(* IEC 61131-3 sources: Jog-the-Robot/plc-for-usb, 2 files *)

(* ---- Main.st ---- *)
(*********************************************************************************
 * Copyright: B&R Industrial Automation GmbH
 * Author:    huebnern
 * Created:   January 23, 2020/8:20 AM
 * Edited:    October 26, 2026 - phone jog, power and home via ESP32 (action RemoteJog)
 *********************************************************************************)
//Main control of the system
PROGRAM _INIT

	//Init Status error
	MainPar.VisuPars.InError 	:= FALSE;
	MainPar.VisuPars.NotInError	:= TRUE;

	//Init Jog velocity
	JogVelocity 				:= INIT_JOG_VELOCITY;

	//Allow jog (Icmp_Ping task is not used)
	AllowJog := TRUE;

	Teach_Pos[0].Pos.X						:=	240;
	Teach_Pos[0].Pos.Y						:= 	0;
	Teach_Pos[0].Pos.Z						:=	335;
	Teach_Pos[0].Orient.Angle1				:=	0;
	Teach_Pos[0].Orient.Angle2				:=	0;

	Teach_Pos[1].Pos.X := 20.699866696484403;
	Teach_Pos[1].Pos.Y := -16.763507571369498;
	Teach_Pos[1].Pos.Z	:= 680.95033173265676;
	Teach_Pos[1].Orient.Angle1 := -126.89365872204304;
	Teach_Pos[1].Orient.Angle2 := 140.99818452000619;

	Teach_Pos[2].Pos.X := -69.244968642624457;
	Teach_Pos[2].Pos.Y := 56.0771029659347;
	Teach_Pos[2].Pos.Z	:= 672.76899259820129;
	Teach_Pos[2].Orient.Angle1 := -111.97058904528618;
	Teach_Pos[2].Orient.Angle2 := 140.99818452000619;

	Teach_Pos[3].Pos.X := 240;
	Teach_Pos[3].Pos.Y := 0;
	Teach_Pos[3].Pos.Z	:= 335;
	Teach_Pos[3].Orient.Angle1 := 0;
	Teach_Pos[3].Orient.Angle2 := 0;

END_PROGRAM

PROGRAM _CYCLIC
	Aktor := Sensor;
	//Error Reset
	fbMpRobotic5Arm.ErrorReset				:= MainPar.Cmd.ErrorReset;

	//Write status
	StatusMain;

	//Change visualization vars
	VisuDisable;

	//Phone jog via ESP32 (BLE -> Modbus TCP). Must run before the state machine.
	RemoteJog;

	//Power On
	IF MainPar.Cmd.PowerOn THEN
		IF fbMpRobotic5Arm.Info.ReadyToPowerOn AND MainPar.StateMachine = STATE_Disabled THEN
			MainPar.StateMachine 	:= STATE_PowerOn;
		END_IF
	ELSE
		MainPar.StateMachine 		:= STATE_Disabled;
	END_IF

	//---------------------------------------------
	//-------------State Machine-------------------
	//---------------------------------------------
	CASE MainPar.StateMachine OF

		//--------State Disabled-------------------
		STATE_Disabled:

			//Power robot off
			fbMpRobotic5Arm.Power 			:= FALSE;

			//Set PreStateIdent
			MainPar.PreStateIdent 			:= STATE_Disabled;

			//Reset Error as long as the robot is disabled
			MainPar.VisuPars.InError 	:= FALSE;
			MainPar.VisuPars.NotInError	:= TRUE;

		//--------State PowerOn-------------------
		STATE_PowerOn:

			//Power robot on
			fbMpRobotic5Arm.Power 			:= TRUE;

			IF MainPar.Status = Idle THEN
				MainPar.StateMachine 		:= STATE_WaitForHome;
			END_IF

		//--------State WaitForHome-------------------
		STATE_WaitForHome:

			//Set PreStateIdent
			MainPar.PreStateIdent 			:= STATE_WaitForHome;

			//Reset Stop
			IF fbMpRobotic5Arm.Stop THEN
				fbMpRobotic5Arm.Stop 		:= FALSE;
			END_IF

			IF MainPar.Cmd.Home THEN
				MainPar.StateMachine 	:= STATE_Home;
				MainPar.HomingCount		:= NoHoming;
				//Reset command
				MainPar.Cmd.Home 		:= FALSE;
			END_IF

		//--------State Home-------------------
		STATE_Home:

			fbMpRobotic5Arm.Home := TRUE;

			IF MainPar.HomingCount = NoHoming THEN
				ChangeHomingMode := FALSE;
			ELSIF MainPar.HomingCount = DefaultHomingDone THEN
				ChangeHomingMode := TRUE;
			END_IF

			IF EDGEPOS(fbMpRobotic5Arm.IsHomed) THEN
				MainPar.HomingCount 		:= MainPar.HomingCount + 1;
				fbMpRobotic5Arm.Home 		:= FALSE;
			END_IF

			IF MainPar.HomingCount = DirectHomingDone THEN
				MainPar.StateMachine 		:= STATE_Idle;
				fbMpRobotic5Arm.Home 		:= FALSE;
			ELSIF MainPar.Cmd.Stop THEN
				MainPar.StateMachine 		:= STATE_WaitForHome;
				fbMpRobotic5Arm.Stop 		:= TRUE;
				fbMpRobotic5Arm.Home 		:= FALSE;
				//Reset command
				MainPar.Cmd.Stop 			:= FALSE;
			END_IF

		//--------State Idle-------------------
		STATE_Idle:

			//Set PreStateIdent
			MainPar.PreStateIdent 			:= STATE_Idle;

			//Reset Stop
			IF fbMpRobotic5Arm.Stop THEN
				fbMpRobotic5Arm.Stop 		:= FALSE;
			END_IF

			IF MainPar.Cmd.Home THEN
				MainPar.HomingCount			:= NoHoming;
				MainPar.StateMachine 		:= STATE_Home;

			ELSE

				//Change to GCode state in case of visu is currently on the G-Code page
				IF (MainPar.GoToState.GCode) AND EDGEPOS(MainPar.Cmd.Start) THEN
					MainPar.StateMachine 	:= STATE_GCode;
				END_IF

				//Change to Tipping state in case of visu is currently on the Tipping page (or the phone has control)
				IF (MainPar.GoToState.Tipping) AND (JogDirectionSet) THEN
					MainPar.StateMachine 	:= STATE_Tipping;
				END_IF

				//Change to MoveSetPos state in case of visu is currently on the MoveSetPos page
				IF (MainPar.GoToState.MoveSetPos) AND EDGEPOS(MainPar.Cmd.Start) THEN
					MainPar.StateMachine 	:= STATE_MoveSetPos;
				END_IF

			END_IF

		//--------State G-Code-------------------
		STATE_GCode:

			//Start movement
			fbMpRobotic5Arm.MoveProgram 		:= TRUE;

			//Stop movement
			IF MainPar.Cmd.Stop THEN
				fbMpRobotic5Arm.Stop 			:= TRUE;
				fbMpRobotic5Arm.MoveProgram 	:= FALSE;
				MainPar.StateMachine 			:= STATE_Idle;
			ELSIF fbMpRobotic5Arm.MoveDone THEN
				fbMpRobotic5Arm.MoveProgram 	:= FALSE;
				MainPar.StateMachine 			:= STATE_Idle;
			END_IF

		//--------State Tipping-------------------
		STATE_Tipping:

			//Change coordinate system
			ParRobot.CoordSystem 			:= mcACS;

			//Set velocity for chosen axis with action
			Tipping;

			//Call Jog
			IF AllowJog THEN
				fbMpRobotic5Arm.Jog := TRUE;
			ELSE
				fbMpRobotic5Arm.Jog := FALSE;
			END_IF

			IF NOT JogDirectionSet THEN
				MainPar.StateMachine 		:= STATE_Idle;
				fbMpRobotic5Arm.Jog 		:= FALSE;
			END_IF

		//--------State MoveSetPos-------------------
		STATE_MoveSetPos:

			//Change coordinate system
			ParRobot.CoordSystem 				:= mcMCS;

			//Start movement
			IF MainPar.Cmd.MoveIndex THEN
				fbMpRobotic5Arm.MoveDirect 	:= TRUE;
			ELSIF NOT MainPar.Cmd.MoveIndex THEN
				fbMpRobotic5Arm.MoveLinear 	:= TRUE;
			END_IF

			//Stop movement
			IF MainPar.Cmd.Stop THEN
				fbMpRobotic5Arm.Stop 			:= TRUE;
				fbMpRobotic5Arm.MoveDirect 	:= FALSE;
				fbMpRobotic5Arm.MoveLinear 	:= FALSE;
				MainPar.StateMachine 			:= STATE_Idle;
			ELSIF fbMpRobotic5Arm.MoveDone THEN
				fbMpRobotic5Arm.MoveDirect 	:= FALSE;
				fbMpRobotic5Arm.MoveLinear 	:= FALSE;
				MainPar.StateMachine 			:= STATE_Idle;
			END_IF

		//--------State Error-------------------
		STATE_Error:

			//Set output var for visu
			MainPar.VisuPars.InError 		:= TRUE;
			MainPar.VisuPars.NotInError		:= FALSE;

			//Stop movement
			fbMpRobotic5Arm.Stop 			:= TRUE;
			fbMpRobotic5Arm.MoveDirect 	:= FALSE;
			fbMpRobotic5Arm.MoveLinear 	:= FALSE;
			fbMpRobotic5Arm.Jog 			:= FALSE;
			fbMpRobotic5Arm.MoveProgram 	:= FALSE;
			fbMpRobotic5Arm.Home 			:= FALSE;

			//Go out of the error state as soon as no error is active
			IF MainPar.Status <> Error THEN
				MainPar.StateMachine 		:= MainPar.PreStateIdent;
				fbMpRobotic5Arm.Stop 		:= FALSE;
				MainPar.VisuPars.InError 	:= FALSE;
				MainPar.VisuPars.NotInError	:= TRUE;
				MainPar.Cmd.ErrorReset		:= FALSE;
			END_IF

	END_CASE

END_PROGRAM

PROGRAM _EXIT

END_PROGRAM

(* ---- RemoteJog.st ---- *)
(*********************************************************************************
 * Action RemoteJog (task Main)  -  version 2: jog + power + home + stop + safety interlocks
 * Lets the Android app control the robot through the ESP32 (BLE -> Modbus TCP).
 * The ESP32 (194.94.86.15) is read and written by the Modbus device "ModbusTcp_any":
 *   read  (FC4):  BleHeartbeat, BleEnable, BleAxis, BleDir, BleCmd, BleCmdSeq
 *   write (FC16): BleStateOut, BleHbEcho
 * Called in Main _CYCLIC right after "VisuDisable;".
 *********************************************************************************)
ACTION RemoteJog:

	// 1. Watchdog: the ESP32 heartbeat must change at least every 500 ms
	IF BleHeartbeat <> BleHeartbeatOld THEN
		BleHeartbeatOld 			:= BleHeartbeat;
		BleWatchdog.IN 				:= FALSE;
	ELSE
		BleWatchdog.IN 				:= TRUE;
	END_IF
	BleWatchdog.PT 					:= T#500ms;
	BleWatchdog();
	BleLinkOk 						:= NOT BleWatchdog.Q;

	// 2. Who has control? The phone takes over while it is connected, but never
	//    in the middle of a running program: then it only watches, and takes
	//    over as soon as the program has ended.
	BleProgramRunning 				:= (MainPar.StateMachine = STATE_GCode) OR (MainPar.StateMachine = STATE_MoveSetPos);

	IF BleLinkOk AND BleEnable = 1 THEN
		IF NOT BleRemoteActive AND NOT BleProgramRunning THEN
			BleRemoteActive 		:= TRUE;
		END_IF
	ELSIF BleRemoteActive THEN
		// Link lost or phone gone: stop and give control back to the panel
		BleRemoteActive 			:= FALSE;
		JogDirection.Positive 		:= FALSE;
		JogDirection.Negative 		:= FALSE;
		MainPar.GoToState.Tipping 	:= FALSE;
	END_IF

	// Fresh press: a jog only counts if the button was pressed while the robot
	// was Ready (or already jogging). A button that was held while a program ran
	// or while homing is ignored until it is released and pressed again.
	IF BleDir = 0 THEN
		BleJogArmed 				:= TRUE;
	ELSIF NOT (MainPar.StateMachine = STATE_Idle OR MainPar.StateMachine = STATE_Tipping) THEN
		BleJogArmed 				:= FALSE;
	END_IF

	// 3. Jog
	IF BleRemoteActive THEN

		// Tells the panel "jog mode": this hides its Start/Stop buttons, so no
		// program can be started while the phone has control.
		MainPar.GoToState.Tipping 	:= TRUE;

		// Select the axis the same way the panel does (ImageIndex ranges ax1..ax5)
		CASE BleAxis OF
			1: IF ImageIndex < ax1 OR ImageIndex > ax1pos THEN ImageIndex := ax1; END_IF
			2: IF ImageIndex < ax2 OR ImageIndex > ax2pos THEN ImageIndex := ax2; END_IF
			3: IF ImageIndex < ax3 OR ImageIndex > ax3pos THEN ImageIndex := ax3; END_IF
			4: IF ImageIndex < ax4 OR ImageIndex > ax4pos THEN ImageIndex := ax4; END_IF
			5: IF ImageIndex < ax5 OR ImageIndex > ax5pos THEN ImageIndex := ax5; END_IF
		END_CASE

		// 1 = positive (R), 2 = negative (L), anything else = stop
		JogDirection.Positive 		:= BleJogArmed AND (BleDir = 1) AND (BleAxis >= 1) AND (BleAxis <= 5);
		JogDirection.Negative 		:= BleJogArmed AND (BleDir = 2) AND (BleAxis >= 1) AND (BleAxis <= 5);

	END_IF

	// 4. Robot commands (power, home). The ESP32 counts BleCmdSeq up by one for
	//    every tap in the app; we act once on every new number.
	IF NOT BleLinkOk THEN
		// After a lost link (or a PLC/ESP32 restart) the first value is only
		// remembered, never executed, so an old command can't run by surprise.
		BleSeqSynced 				:= FALSE;
	ELSIF NOT BleSeqSynced THEN
		BleCmdSeqOld 				:= BleCmdSeq;
		BleSeqSynced 				:= TRUE;
	ELSIF BleCmdSeq <> BleCmdSeqOld THEN
		BleCmdSeqOld 				:= BleCmdSeq;
		CASE BleCmd OF
			1: // Power on
				MainPar.Cmd.PowerOn := TRUE;
			2: // Power off, but never while the robot is moving
				IF NOT (BleProgramRunning OR MainPar.StateMachine = STATE_Tipping OR MainPar.StateMachine = STATE_Home) THEN
					MainPar.Cmd.PowerOn := FALSE;
					BleHomeRequest 	:= FALSE;
				END_IF
			3: // Home, only when the robot can home
				IF MainPar.StateMachine = STATE_WaitForHome OR MainPar.StateMachine = STATE_Idle THEN
					BleHomeRequest 	:= TRUE;
				END_IF
			4: // Stop a running program, move or homing
				IF BleProgramRunning OR MainPar.StateMachine = STATE_Home THEN
					BleStopRequest 	:= TRUE;
				END_IF
		END_CASE
	END_IF

	// Stop works like the panel's Stop push button: Cmd.Stop stays TRUE until
	// the state machine has left the program/move/homing state, then it is
	// released. Once the robot is Ready again, the phone takes control (step 2).
	IF BleStopRequest THEN
		IF BleProgramRunning OR MainPar.StateMachine = STATE_Home THEN
			MainPar.Cmd.Stop 		:= TRUE;
		ELSE
			MainPar.Cmd.Stop 		:= FALSE;
			BleStopRequest 			:= FALSE;
		END_IF
	END_IF

	// Home works like the panel's push button: Cmd.Home stays TRUE until the
	// state machine has entered STATE_Home, then it is released again.
	IF BleHomeRequest THEN
		IF MainPar.StateMachine = STATE_Home OR MainPar.StateMachine = STATE_Disabled THEN
			MainPar.Cmd.Home 		:= FALSE;
			BleHomeRequest 			:= FALSE;
		ELSE
			MainPar.Cmd.Home 		:= TRUE;
		END_IF
	END_IF

	// 5. Feedback to the ESP32 (and from there to the app)
	CASE MainPar.StateMachine OF
		STATE_Disabled:		BleStateOut := 0;
		STATE_PowerOn:		BleStateOut := 5;
		STATE_WaitForHome:	BleStateOut := 9;
		STATE_Home:			BleStateOut := 10;
		STATE_Idle:			BleStateOut := 20;
		STATE_GCode:		BleStateOut := 30;
		STATE_Tipping:		BleStateOut := 40;
		STATE_MoveSetPos:	BleStateOut := 50;
		STATE_Error:		BleStateOut := 99;
	END_CASE
	BleHbEcho 						:= BleHeartbeat;	// proves to the ESP32 that the PLC is running

END_ACTION
